// TwinCAT 3 PLC project ModeOutputsTests
// ProgramVersion: 3.1.4026.22
// libraries:
//   Tc2_Standard, * (Beckhoff Automation GmbH)
//   Tc2_System, * (Beckhoff Automation GmbH)
// project tree:
//   StateMachineControl/DUTs/ E_ModeState.TcDUT, ST_ModeOutputs.TcDUT
//   StateMachineControl/GVLs/ GVL_MODE.TcGVL
//   StateMachineControl/POUs/ F_DeriveModeOutputs.TcPOU
//   StateMachineControl/tests/POUs/ PRG_ModeOutputsTests.TcPOU
//   StateMachineControl/tests/ ModeOutputsTestTask.TcTTO
// (motion and I/O tree: see PLC project experimentsequencertests)
// real-time tasks:
//   TASK DriveStateTestTask: cycle T#10ms, priority 1, ADS port 350
//   TASK TestTask: cycle T#10ms, priority 2, ADS port 351

CONFIGURATION ModeOutputsTests
    RESOURCE PLC ON TwinCAT3
        TASK ModeOutputsTestTask(INTERVAL := T#10ms, PRIORITY := 1);
        PROGRAM PRG_ModeOutputsTests WITH ModeOutputsTestTask : PRG_ModeOutputsTests;
    END_RESOURCE
END_CONFIGURATION

// ---- StateMachineControl/DUTs/E_ModeState.TcDUT
{attribute 'qualified_only'}
{attribute 'strict'}
{attribute 'to_string'}
TYPE E_ModeState :
(
    IDLE := 0,              // Servo OFF / initial
    RESETTING := 10,        // Reset pulse active — no experiment transitions allowed
    SERVO_READY := 20,      // Servo ON + drive OPERATION_ENABLED, awaiting experiment
    RUNNING := 30,          // Experiment active
    DONE := 40              // Playback complete, awaiting rearm
);
END_TYPE

// ---- StateMachineControl/DUTs/ST_ModeOutputs.TcDUT
TYPE ST_ModeOutputs :
STRUCT
    experimentActiveOut : BOOL;
    preArmOut : BOOL;
    resetOut : BOOL;
    enableCurrentOut : BOOL;
END_STRUCT
END_TYPE

// ---- StateMachineControl/GVLs/GVL_MODE.TcGVL
{attribute 'qualified_only'}
VAR_GLOBAL CONSTANT
    MODEF_SERVO_ENABLE : UINT := 16#0001;          (* bit0 *)
    MODEF_EXPERIMENT_START_REQ : UINT := 16#0002;  (* bit1 *)
    HEARTBEAT_TIMEOUT_TICKS : UDINT := 50;         (* 10 ms task * 50 = 500 ms *)

END_VAR

VAR_GLOBAL
    {attribute 'linkalways'}
    modeFlags : UINT := 0;
    resetReq : BOOL := FALSE;
    resetAckCounter : UDINT := 0;
    hostHeartbeatCounter : UDINT := 0;
    watchdogTripCounter : UDINT := 0;
    experimentActive : BOOL := FALSE;
    loggerFileReleased : BOOL := FALSE;
    loggerErrorCode : UDINT := 0;
    modeState : E_ModeState := E_ModeState.IDLE;
END_VAR

// ---- StateMachineControl/tests/POUs/PRG_ModeOutputsTests.TcPOU
PROGRAM PRG_ModeOutputsTests
VAR
    outputs : ST_ModeOutputs;
    testsExecuted : BOOL := FALSE;
    testsPassed : BOOL := FALSE;
    failureCount : UDINT := 0;
END_VAR

IF NOT testsExecuted THEN
    outputs := F_DeriveModeOutputs(modeState := E_ModeState.IDLE);
    IF outputs.experimentActiveOut OR outputs.preArmOut OR outputs.resetOut
        OR outputs.enableCurrentOut THEN
        failureCount := failureCount + 1;
    END_IF

    outputs := F_DeriveModeOutputs(modeState := E_ModeState.RESETTING);
    IF outputs.experimentActiveOut OR outputs.preArmOut OR NOT outputs.resetOut
        OR outputs.enableCurrentOut THEN
        failureCount := failureCount + 1;
    END_IF

    outputs := F_DeriveModeOutputs(modeState := E_ModeState.SERVO_READY);
    IF outputs.experimentActiveOut OR NOT outputs.preArmOut OR outputs.resetOut
        OR NOT outputs.enableCurrentOut THEN
        failureCount := failureCount + 1;
    END_IF

    outputs := F_DeriveModeOutputs(modeState := E_ModeState.RUNNING);
    IF NOT outputs.experimentActiveOut OR outputs.preArmOut OR outputs.resetOut
        OR NOT outputs.enableCurrentOut THEN
        failureCount := failureCount + 1;
    END_IF

    outputs := F_DeriveModeOutputs(modeState := E_ModeState.DONE);
    IF outputs.experimentActiveOut OR outputs.preArmOut OR outputs.resetOut
        OR outputs.enableCurrentOut THEN
        failureCount := failureCount + 1;
    END_IF

    (* Consecutive calls must not retain fields from the previous state. *)
    outputs := F_DeriveModeOutputs(modeState := E_ModeState.RUNNING);
    outputs := F_DeriveModeOutputs(modeState := E_ModeState.IDLE);
    IF outputs.experimentActiveOut OR outputs.preArmOut OR outputs.resetOut
        OR outputs.enableCurrentOut THEN
        failureCount := failureCount + 1;
    END_IF

    testsExecuted := TRUE;
    testsPassed := (failureCount = 0);
END_IF

END_PROGRAM

// ---- StateMachineControl/POUs/F_DeriveModeOutputs.TcPOU
FUNCTION F_DeriveModeOutputs : ST_ModeOutputs
VAR_INPUT
    modeState : E_ModeState;
END_VAR

(* Safe default for unknown or newly added states. *)
F_DeriveModeOutputs.experimentActiveOut := FALSE;
F_DeriveModeOutputs.preArmOut := FALSE;
F_DeriveModeOutputs.resetOut := FALSE;
F_DeriveModeOutputs.enableCurrentOut := FALSE;

CASE modeState OF
    E_ModeState.RESETTING:
        F_DeriveModeOutputs.resetOut := TRUE;

    E_ModeState.SERVO_READY:
        F_DeriveModeOutputs.preArmOut := TRUE;
        F_DeriveModeOutputs.enableCurrentOut := TRUE;

    E_ModeState.RUNNING:
        F_DeriveModeOutputs.experimentActiveOut := TRUE;
        F_DeriveModeOutputs.enableCurrentOut := TRUE;
END_CASE

END_FUNCTION
